Staubli VAL3: teachPoint.pgx

program teachPoint(num x_nIndex)
  local bool l_bResult
  local pointRx l_pPoint
  local tool l_tTool
begin
  l_bResult=userPageConfirm("是否记录当前点位？")
  if l_bResult
    call saveData:getTool(saveData:nJogTool,l_tTool)
    fFrame.trsf.x=nFrame[0]
    fFrame.trsf.y=nFrame[1]
    fFrame.trsf.z=nFrame[2]
    fFrame.trsf.rx=nFrame[3]
    fFrame.trsf.ry=nFrame[4]
    fFrame.trsf.rz=nFrame[5]

    l_pPoint=here(l_tTool,fFrame)
    safeTemp:zZoneItem[x_nIndex].pFirst.trsf=l_pPoint.trsf
    safeTemp:zZoneItem[x_nIndex].pFirst.config=l_pPoint.config
    safeTemp:libSave()




    delay(0.1)
  endIf
end
